(* IEC 61131-3 sources: nautilus/siemens/writer/testdata/tasks, 4 files *)

(* ---- types.st ---- *)
(* The project's library: the struct a shared tag is. *)
TYPE
  Motor : STRUCT
    Run   : BOOL;
    Speed : REAL;
  END_STRUCT;
END_TYPE

(* ---- Fast.st ---- *)
(* A faster task: writes one shared tag, and reads tags the main task
   writes through a timer's and a latch's output bindings. *)
PROGRAM Fast
VAR_EXTERNAL
  Pump : Motor;
  Level : REAL;
END_VAR
IF Pump.Run AND NOT (Done OR Alarm) THEN
  Level := Level + Pump.Speed * 0.01;
ELSE
  Level := Level - 0.5;
END_IF;
END_PROGRAM

(* ---- Main.st ---- *)
(* The main task: a seal-in on a shared tag (assigned every scan, often
   to the value it has), a struct member, a timer output and a latch bound
   to shared tags, a tag no other task names, and a RETURN. *)
PROGRAM Main
VAR_EXTERNAL
  Start : BOOL;
  Stop : BOOL;
  Run : BOOL;
  Pump : Motor;
  Level : REAL;
  Done : BOOL;
  Alarm : BOOL;
  Status : WORD;
  Local1 : DINT;
END_VAR
VAR
  dwell : TON;
  latch : SR;
  Name : INT;
END_VAR
Run := (Start OR Run) AND NOT Stop;
Pump.Run := Run AND Level < 90.0;
dwell(IN := Run, PT := T#5s, Q => Done);
latch(S1 := Level > 95.0, R := Stop, Q1 => Alarm);
Local1 := Local1 + 1;
Name := Name + 1;
IF NOT Status.3 THEN
  RETURN;
END_IF;
Pump.Speed := 0.0;
END_PROGRAM

(* ---- Slow.st ---- *)
(* A slower task: writes single bits of a shared word and, sometimes,
   the whole word; and names its tags with no VAR_EXTERNAL (implicit
   scope). *)
PROGRAM Slow
VAR
  i : INT;
END_VAR
Status.3 := Level > 10.0;
IF Stop THEN
  Status.0 := TRUE;
END_IF;
IF Start THEN
  Status := 16#0;
END_IF;
FOR i := 1 TO 3 DO
  Status.7 := NOT Status.7;
END_FOR;
END_PROGRAM
